// TIA Portal V20 export
// export: Created 2026-10-12T04:58:21.9485883Z, ExportSetting WithDefaults, DisplayName Totally Integrated Automation Portal, DisplayVersion V20, DisplayName TIA Portal Openness, DisplayVersion V20, DisplayName TIA Portal Teamcenter Gateway, DisplayVersion V20, DisplayName TIA Portal Version Control Interface, DisplayVersion V20, DisplayName SINAMICS Startdrive Advanced, DisplayVersion V20 SP1 Update 2, DisplayName SINAMICS Startdrive G110M, G120, G120C, G120D, G120P, G115D, DisplayVersion V20 SP1 Update 2, DisplayName SINAMICS Startdrive G130, G150, S120, S150, SINAMICS MV, G220, S200, S210, DisplayVersion V20 SP1 Update 2, DisplayName STEP 7 Professional, DisplayVersion V20, DisplayName STEP 7 Safety, DisplayVersion V20, DisplayName WinCC Basic/Comfort/Advanced, DisplayVersion V20, DisplayName WinCC Professional, DisplayVersion V20, DisplayName WinCC Unified, DisplayVersion V20
FUNCTION "FRK_SetBoot" : Void   // FC117, SCL
{ S7_Optimized_Access := 'TRUE' }
VERSION : 0.1
// stored: AutoNumber true, IsIECCheckEnabled false, SetENOAutomatically false, UDAEnableTagReadback false
   VAR_INPUT
      Startup : Bool;
   END_VAR
   VAR_TEMP
      RootIndex : Int;
      Slot : Int;
   END_VAR
BEGIN

   IF NOT #Startup THEN
       RETURN;
   END_IF;
   IF "FRK_SetStore".SchemaVersion <> 1 THEN
       FOR #RootIndex := 1 TO 2 DO
           IF "FRK_SetStore".SchemaVersion <> 0 THEN
               "FRK_ConfigLoss"(RootIndex := #RootIndex,
                                Scope := "FRK_SetStore".Sets[#RootIndex, 1].Info.RootIdentity);
           END_IF;
           FOR #Slot := 1 TO 4 DO
               "FRK_SetStore".Sets[#RootIndex, #Slot].Info.Used := FALSE;
           END_FOR;
       END_FOR;
       "FRK_SetStore".SchemaVersion := 1;
   END_IF;
END_FUNCTION
